FUNCTION_BLOCK FB_Axis EXTENDS FB_Device IMPLEMENTS I_SpeedController
VAR_INPUT
	localEnable		: BOOL; // Enable signal from local Estops, etc. If parent control is configured for enable with no local enable, this can be latched true
	
	{attribute 'OPC.UA.DA' := '1'}
	{attribute 'OPC.UA.DA.StructuredType' := '1'}
	cfg				: ST_AxisConfiguration; 
	
	{attribute 'OPC.UA.DA' := '1'}
	{attribute 'OPC.UA.DA.StructuredType' := '1'}
	ctrlAxis		: ST_AxisControl;
	
	{attribute 'OPC.UA.DA' := '1'} 
	ocmd			: E_AxisCommand;
	
	func			: ST_AxisFunctions;
	
	(* Interlocks/Permissives
	----------------------------------------------------------------------------------------------------*)
	{attribute 'OPC.UA.DA' := '1'}
	{attribute 'OPC.UA.DA.Access' := '1'}
	fwdIntlk		: FB_Permissive;	
	{attribute 'OPC.UA.DA' := '1'}
	{attribute 'OPC.UA.DA.Access' := '1'}
	fwdPerm			: FB_Permissive; 
	{attribute 'OPC.UA.DA' := '1'}
	{attribute 'OPC.UA.DA.Access' := '1'}
	revIntlk		: FB_Permissive; 
	{attribute 'OPC.UA.DA' := '1'}
	{attribute 'OPC.UA.DA.Access' := '1'}
	revPerm			: FB_Permissive; 
	
	(* External inputs
	----------------------------------------------------------------------------------------------------*)
	inpHomeProx AT %I* : BOOL; 				// Link this to home sensor in MapInputs method of Parent
	driveDiagnosticNumber AT %I* : UDINT;	// Link to AX5000 S-0-0390 Diagnostic number
	inpFault		   : BOOL;
	inpFaultText	   : T_MaxString;
END_VAR

VAR_OUTPUT
	{attribute 'OPC.UA.DA' := '1'}
	{attribute 'OPC.UA.DA.StructuredType' := '1'}
	motionParam	: ST_AxisMotionParameters;
	
	{attribute 'OPC.UA.DA' := '1'}
	{attribute 'OPC.UA.DA.Access' := '1'}
	{attribute 'OPC.UA.DA.StructuredType' := '1'}
	sts			: ST_AxisDeviceStatus; 

	{attribute 'OPC.UA.DA' := '1'}
	{attribute 'OPC.UA.DA.Access' := '1'}
	{attribute 'OPC.UA.DA.StructuredType' := '1'}	
	fault		: ST_AxisFault;
END_VAR

VAR PERSISTENT
	offset			: LREAL; // Offset for zero position
	
	{attribute 'OPC.UA.DA' := '1'}
	{attribute 'OPC.UA.DA.Access' := '1'}
	{attribute 'OPC.UA.DA.StructuredType' := '1'}
	positionList	: ARRAY[0..GVL_Lib_ServoConstants.MAX_POSITIONS] OF ST_AxisPosition;
END_VAR

VAR
	axis					: AXIS_REF; 			 // Linked to Motion Axis Object	
	mc						: ST_AxisMotionControl;  // Motion Commands and Parameters
	saveData				: FB_WritePersistentData;
	savePositionListData	: BOOL;	
	resetErrorAndDrive		: BOOL;	
	safeDisable				: BOOL;					 // Disable drive after a safe command, must reset errors to resume operation	
	homingInProgress		: BOOL;					 // Internal bit to set complete flag after homing offset is stored
	mcGearIn				: MC_GearIn;
	mcGearOut				: MC_GearOut;
	
	(* State
	----------------------------------------------------------------------------------------------------*)
	lastGoodState			: E_AxisState;
	nextState				: E_AxisState;
	lastFaultId				: UDINT;
	
	(* Servo Commands
	----------------------------------------------------------------------------------------------------*)
	cmdReceived				: E_AxisCommand;	
	cmdReceivedLast			: E_AxisCommand;	
	pcmd					: E_AxisCommand;	
	pcmdLast				: E_AxisCommand;	
	ocmdLast				: E_AxisCommand;
	storedRelMovePosition	: LREAL;	
	
	(* Speed history/triggers
	----------------------------------------------------------------------------------------------------*)
	jogSpeedLast			: LREAL; 	
	jogSpeedChanged			: BOOL; 	// Jog speed has changed
	ftJogSpeedChanged		: F_TRIG;
	moveSpeedLast			: LREAL;
	moveSpeedChanged		: BOOL;		// Move speed has changed
	ftMoveSpeedChanged		: F_TRIG;
	ftRelMove				: F_TRIG;
	rtAbsMoveADone			: R_TRIG;
	rtAbsMoveBDone			: R_TRIG;
	rtModMoveADone			: R_TRIG;
	rtModMoveBDone			: R_TRIG;

	(* General
	----------------------------------------------------------------------------------------------------*)	
	enableAxisDelay			: TON;
	mcPowerTimeout			: TON;
END_VAR

SUPER^();

Device();
Hmi();
StatusIn();
ProcessCommands();
StateMachine();
MotionControl();
HandleFaults();
StatusOut();
Functions();
SetPositionIds();

METHOD PUBLIC AbsMove
VAR_INPUT
	absMovePosition		: LREAL;
END_VAR
SetMotionParam(param := E_MotorMotionParam.AbsMovePosition, val := absMovePosition);
pcmd := E_AxisCommand.AbsMove;
END_METHOD

METHOD PUBLIC AbsMoveToStoredPosition : BOOL
// Returns true if position is found in list and move started, false otherwise
VAR_INPUT
	id				: INT; 
END_VAR
VAR
	i				: INT;
	success			: BOOL := FALSE;
END_VAR
// Loop through position list to check if the position ID exists and initiate move
FOR i := 0 TO GVL_Lib_ServoConstants.MAX_POSITIONS DO
	// If ID exists in position list
	IF positionList[i].id = id THEN 
		SetMotionParam(param := E_MotorMotionParam.AbsMovePositionId, val := id); // Store commanded position ID
		AbsMove(positionList[i].position); 										  // Initiate absolute move
		success := TRUE;
		EXIT;
	END_IF
END_FOR

AbsMoveToStoredPosition := success;
END_METHOD

METHOD PUBLIC AddFollower
// Must continuously call function
// Execution of coupling or decoupling will be set by 
// the ctrlAxis.coupleFollower bit
VAR_IN_OUT
	follower : AXIS_REF;
END_VAR
IF __ISVALIDREF(follower) THEN
	mcGearIn(Master := axis, Slave := follower, RatioNumerator := cfg.gearRatio, RatioDenominator := 1); 
	mcGearOut(Slave := follower); 

	IF axis.status.homed AND follower.status.homed AND ctrlAxis.coupleFollower
	AND NOT mcGearIn.InGear AND NOT mcGearIn.Execute THEN
		mcGearIn.Execute := TRUE; 
	END_IF

	IF mcGearIn.Execute AND follower.status.coupled THEN 
		mcGearIn.Execute 		:= FALSE;
		ctrlAxis.coupleFollower := TRUE;
	END_IF

	IF mcGearIn.Error THEN
		mcGearIn.Execute := FALSE;
	END_IF

	IF NOT ctrlAxis.coupleFollower AND follower.Status.Coupled THEN 
		mcGearOut.Execute := TRUE;
	END_IF

	IF mcGearOut.Done THEN 
		mcGearOut.Execute := FALSE;
	END_IF

	fault.coupleError 		:= ctrlAxis.coupleFollower AND (NOT axis.Status.Homed OR NOT follower.Status.Homed);
	fault.followerLagError 	:= ctrlAxis.coupleFollower AND axis.Status.Coupled AND follower.Status.Coupled AND
						  	   ABS(axis.NcToPlc.PosDiff - follower.NcToPlc.PosDiff) > cfg.followerLag;			   
END_IF
END_METHOD

METHOD PUBLIC DefinePosition : INT // Check for blank name before overwriting
VAR_INPUT
	id					: INT; // position id
	position			: LREAL; // value of position (mm)
	name				: STRING := ''; // position name
END_VAR
IF positionList[id].name = '' THEN
	DefinePosition := SavePosition(id := id, position := position, name := name);
ELSE
	DefinePosition := 2; // Position has previously been defined. don't overwrite
END_IF
END_METHOD

METHOD PUBLIC DeletePosition : INT
VAR_INPUT
	id : INT;
END_VAR
IF id >= 0 AND id <= GVL_Lib_ServoConstants.MAX_POSITIONS THEN
	positionList[id].name := '';
	positionList[id].position := 0.0;
	DeletePosition := 1; //position deleted, code = 1
ELSE
	DeletePosition := -1; //id out of bounds, code = -1
END_IF
END_METHOD

METHOD PROTECTED Device : BOOL
VAR_INPUT
END_VAR
// to FB device
opTimeout  			 := cfg.opTimeout;
opTimeoutEnable 	 := cfg.opTimeoutEnable;
opActivity 			 := ocmd <> E_AxisCommand.None;

// from FB device
sts.mode	   		 := mode;
sts.modeAuto   		 := sts.mode = E_SystemMode.Auto;
sts.modeManual 		 := sts.mode = E_SystemMode.Manual;
sts.manualOvrde		 := ctrl.manualOvrde; 	
sts.bypass 	   		 := ctrl.bypass;		
sts.sim		   		 := ctrl.sim;			
sts.parentConfigured := parentConfigured;
END_METHOD

METHOD DisableCouple : BOOL
VAR_INPUT
END_VAR
ctrlAxis.coupleFollower := FALSE;
END_METHOD

METHOD PUBLIC DisableLag
pcmd := E_AxisCommand.DisableLag;
END_METHOD

METHOD EnableCouple : BOOL
VAR_INPUT
END_VAR
ctrlAxis.coupleFollower := TRUE;
END_METHOD

METHOD PUBLIC EnableLag
pcmd := E_AxisCommand.EnableLag;
END_METHOD

METHOD PROTECTED Functions
VAR
	i 				: INT;
END_VAR
(* Default function FB calls
----------------------------------------------------------------------------------------------------*)
func.AbsMove(				 	hmiTextStatic := CONCAT(cfg.motorId, ' absolute move'));
func.AbsMoveToStoredPosition(	hmiTextStatic := CONCAT(cfg.motorId, ' absolute move to stored position'));
func.RelMove(					hmiTextStatic := CONCAT(cfg.motorId, ' relative move'));
func.ModMove(				 	hmiTextStatic := CONCAT(cfg.motorId, ' modulus move'));
func.LatchJogFwd(			 	hmiTextStatic := CONCAT(cfg.motorId, ' latch jog forward'));
func.LatchJogRev(				hmiTextStatic := CONCAT(cfg.motorId, ' latch jog reverse'));
func.Home(						hmiTextStatic := CONCAT(cfg.motorId, ' home'));
func.Stop(						hmiTextStatic := CONCAT(cfg.motorId, ' stop'));
func.Couple(					hmiTextStatic := CONCAT(cfg.motorId, ' coupling follower'));
func.Decouple(					hmiTextStatic := CONCAT(cfg.motorId, ' decoupling follower'));
func.ResetDoneBits(				hmiTextStatic := CONCAT(cfg.motorId, ' reset done bits'));

(* Default functions
----------------------------------------------------------------------------------------------------*)

IF func.AbsMove.entry THEN
	FOR i := GVL_Lib_SequencerConstants.MIN_PARAMETERS TO GVL_Lib_SequencerConstants.MAX_PARAMETERS DO
		CASE func.AbsMove.arrParam[i].typeEnum OF
			E_AxisFunctionParam.AbsMovePosition:
				SetMotionParam(param	:= E_MotorMotionParam.AbsMovePosition,
							   val		:= func.AbsMove.arrParam[i].value);
			E_AxisFunctionParam.MoveSpeed:
				SetMotionParam(param	:= E_MotorMotionParam.MoveSpeed,
							   val		:= func.AbsMove.arrParam[i].value);
		END_CASE
	END_FOR
END_IF
IF func.AbsMove.running THEN
	// Check for speed change mid move
	FOR i := GVL_Lib_SequencerConstants.MIN_PARAMETERS TO GVL_Lib_SequencerConstants.MAX_PARAMETERS DO
		IF func.AbsMove.arrParam[i].typeEnum = E_AxisFunctionParam.MoveSpeed THEN
			SetMotionParam(param	:= E_MotorMotionParam.MoveSpeed,
						   val		:= func.AbsMove.arrParam[i].value);
		END_IF
	END_FOR
	// Wait for complete conditions
	func.AbsMove.permComplete.perm.0 S= sts.absMoveComplete;
	
	// Call Action
	IF NOT func.AbsMove.complete AND NOT fault.active
	AND sts.state <> E_AxisState.AbsMove_A AND sts.state <> E_AxisState.AbsMove_B THEN
		// Passing in this motion parameter has the effect of reassigning its own 
		// value to itself. It's done because this input is required for the method
		AbsMove(motionParam.absMovePosition);
	END_IF
	
	func.AbsMove.inpError := fault.active;
END_IF


IF func.AbsMoveToStoredPosition.entry THEN
	FOR i := GVL_Lib_SequencerConstants.MIN_PARAMETERS TO GVL_Lib_SequencerConstants.MAX_PARAMETERS DO
		CASE func.AbsMoveToStoredPosition.arrParam[i].typeEnum OF
			E_AxisFunctionParam.AbsMovePositionId:
				SetMotionParam(param	:= E_MotorMotionParam.AbsMovePositionId,
							   val		:= func.AbsMoveToStoredPosition.arrParam[i].value);
			E_AxisFunctionParam.MoveSpeed:
				SetMotionParam(param	:= E_MotorMotionParam.MoveSpeed,
							   val		:= func.AbsMoveToStoredPosition.arrParam[i].value);
		END_CASE
	END_FOR
END_IF
IF func.AbsMoveToStoredPosition.running THEN
	// Check for speed change mid move
	FOR i := GVL_Lib_SequencerConstants.MIN_PARAMETERS TO GVL_Lib_SequencerConstants.MAX_PARAMETERS DO
		IF func.AbsMoveToStoredPosition.arrParam[i].typeEnum = E_AxisFunctionParam.MoveSpeed THEN
			SetMotionParam(param	:= E_MotorMotionParam.MoveSpeed,
						   val		:= func.AbsMoveToStoredPosition.arrParam[i].value);
		END_IF
	END_FOR
	// Wait for complete conditions
	func.AbsMoveToStoredPosition.permComplete.perm.0 S= sts.absMoveComplete;	
	
	// Call Action
	IF NOT func.AbsMoveToStoredPosition.complete AND NOT fault.active
	AND sts.state <> E_AxisState.AbsMove_A AND sts.state <> E_AxisState.AbsMove_B THEN
		AbsMoveToStoredPosition(motionParam.absMovePositionId);
	END_IF
	
	func.AbsMoveToStoredPosition.inpError := fault.active;
END_IF


IF func.RelMove.entry THEN
	FOR i := GVL_Lib_SequencerConstants.MIN_PARAMETERS TO GVL_Lib_SequencerConstants.MAX_PARAMETERS DO
		CASE func.RelMove.arrParam[i].typeEnum OF
			E_AxisFunctionParam.RelMoveDistance:
				SetMotionParam(param	:= E_MotorMotionParam.RelMoveDistance,
							   val		:= func.RelMove.arrParam[i].value);
			E_AxisFunctionParam.MoveSpeed:
				SetMotionParam(param	:= E_MotorMotionParam.MoveSpeed,
							   val		:= func.RelMove.arrParam[i].value);
		END_CASE
	END_FOR
END_IF
IF func.RelMove.running THEN
	// Check for speed change mid move
	FOR i := GVL_Lib_SequencerConstants.MIN_PARAMETERS TO GVL_Lib_SequencerConstants.MAX_PARAMETERS DO
		IF func.RelMove.arrParam[i].typeEnum = E_AxisFunctionParam.MoveSpeed THEN
			SetMotionParam(param	:= E_MotorMotionParam.MoveSpeed,
						   val		:= func.RelMove.arrParam[i].value);
		END_IF
	END_FOR
	// Wait for complete conditions
	func.RelMove.permComplete.perm.0 S= sts.RelMoveComplete;
	
	// Call Action
	IF NOT func.RelMove.complete AND NOT fault.active
	AND sts.state <> E_AxisState.RelMove_A AND sts.state <> E_AxisState.RelMove_B THEN
		RelMove(motionParam.relMoveDistance);
	END_IF
	
	func.RelMove.inpError := fault.active;
END_IF


IF func.ModMove.entry THEN
	FOR i := GVL_Lib_SequencerConstants.MIN_PARAMETERS TO GVL_Lib_SequencerConstants.MAX_PARAMETERS DO
		CASE func.ModMove.arrParam[i].typeEnum OF
			E_AxisFunctionParam.ModMovePosition:
				SetMotionParam(param	:= E_MotorMotionParam.ModMovePosition,
							   val		:= func.ModMove.arrParam[i].value);
			E_AxisFunctionParam.MoveSpeed:
				SetMotionParam(param	:= E_MotorMotionParam.MoveSpeed,
							   val		:= func.ModMove.arrParam[i].value);
		END_CASE
	END_FOR
	END_IF
IF func.ModMove.running THEN
	// Check for speed change mid move
	FOR i := GVL_Lib_SequencerConstants.MIN_PARAMETERS TO GVL_Lib_SequencerConstants.MAX_PARAMETERS DO
		IF func.ModMove.arrParam[i].typeEnum = E_AxisFunctionParam.MoveSpeed THEN
			SetMotionParam(param	:= E_MotorMotionParam.MoveSpeed,
						   val		:= func.ModMove.arrParam[i].value);
		END_IF
	END_FOR
	// Wait for complete conditions
	func.ModMove.permComplete.perm.0 S= sts.ModMoveComplete;
	
	// Call Action
	IF NOT func.ModMove.complete AND NOT fault.active
	AND sts.state <> E_AxisState.ModMove_A AND sts.state <> E_AxisState.ModMove_B THEN
		ModMove(motionParam.modMovePosition);
	END_IF

	func.ModMove.inpError := fault.active;
END_IF


IF func.LatchJogFwd.entry THEN
	FOR i := GVL_Lib_SequencerConstants.MIN_PARAMETERS TO GVL_Lib_SequencerConstants.MAX_PARAMETERS DO
		CASE func.LatchJogFwd.arrParam[i].typeEnum OF
			E_AxisFunctionParam.JogSpeed: 
				SetMotionParam(param	:= E_MotorMotionParam.JogSpeed,
							   val		:= func.LatchJogFwd.arrParam[i].value);
		END_CASE
	END_FOR
END_IF
IF func.LatchJogFwd.running THEN
	// Check for speed change mid move
	FOR i := GVL_Lib_SequencerConstants.MIN_PARAMETERS TO GVL_Lib_SequencerConstants.MAX_PARAMETERS DO
		IF func.LatchJogFwd.arrParam[i].typeEnum = E_AxisFunctionParam.JogSpeed THEN
			SetMotionParam(param	:= E_MotorMotionParam.JogSpeed,
						   val		:= func.LatchJogFwd.arrParam[i].value);
		END_IF
	END_FOR	
	// Call Action
	IF NOT fault.active THEN
		LatchJogFwd();
	END_IF
	
	// Wait for complete conditions
	func.LatchJogFwd.permComplete.perm.0 S= sts.jogFwdInProgress;
	
	func.LatchJogFwd.inpError := fault.active;
END_IF


IF func.LatchJogRev.entry THEN
	FOR i := GVL_Lib_SequencerConstants.MIN_PARAMETERS TO GVL_Lib_SequencerConstants.MAX_PARAMETERS DO
		CASE func.LatchJogRev.arrParam[i].typeEnum OF
			E_AxisFunctionParam.JogSpeed:
				SetMotionParam(param	:= E_MotorMotionParam.JogSpeed,
							   val		:= func.LatchJogRev.arrParam[i].value);
		END_CASE
	END_FOR
END_IF
IF func.LatchJogRev.running THEN
	// Check for speed change mid move
	FOR i := GVL_Lib_SequencerConstants.MIN_PARAMETERS TO GVL_Lib_SequencerConstants.MAX_PARAMETERS DO
		IF func.LatchJogRev.arrParam[i].typeEnum = E_AxisFunctionParam.JogSpeed THEN
			SetMotionParam(param	:= E_MotorMotionParam.JogSpeed,
						   val		:= func.LatchJogRev.arrParam[i].value);
		END_IF
	END_FOR	
	// Call Action
	IF NOT fault.active THEN
		LatchJogRev();
	END_IF
	
	// Wait for complete conditions
	func.LatchJogRev.permComplete.perm.0 S= sts.jogRevInProgress;
	
	func.LatchJogRev.inpError := fault.active;
END_IF



IF func.Home.entry THEN
	FOR i := GVL_Lib_SequencerConstants.MIN_PARAMETERS TO GVL_Lib_SequencerConstants.MAX_PARAMETERS DO
		CASE func.Home.arrParam[i].typeEnum OF
			E_AxisFunctionParam.HomePosition:
				SetMotionParam(param	:= E_MotorMotionParam.HomePosition,
							   val		:= func.Home.arrParam[i].value);
		END_CASE
	END_FOR
END_IF
IF func.Home.running THEN
	// Wait for complete conditions
	func.Home.permComplete.perm.0 S= sts.homingComplete OR ctrl.sim;
	
	// Call Action
	IF NOT func.Home.complete AND NOT fault.active
	AND sts.state <> E_AxisState.Homing THEN
		Home();
	END_IF
	
	func.Home.inpError := fault.active;
END_IF

IF func.Stop.running THEN
	// Wait for complete conditions	
	func.Stop.permComplete.perm.0 S= sts.stopComplete;
	
	// Call action
	IF NOT func.Stop.complete AND NOT fault.active
	AND sts.state <> E_AxisState.Halting THEN
		Stop();
	END_IF
END_IF


IF func.Couple.running THEN
	ctrlAxis.coupleFollower := TRUE;
	func.Couple.PermComplete.perm.0 := sts.coupled;
END_IF


IF func.Decouple.running THEN
	ctrlAxis.coupleFollower := FALSE;
	func.Decouple.PermComplete.perm.0 := NOT sts.coupled;
END_IF


IF func.ResetDoneBits.running THEN
	ctrlAxis.resetDoneBits := TRUE;
	func.ResetDoneBits.permComplete.perm.0 := TRUE;
END_IF
END_METHOD

METHOD PROTECTED HandleFaults : BOOL
VAR
	i					: INT;
END_VAR
(* ----- Set Faults ----- *)
// Axis Drive Device Error
IF axis.Status.DriveDeviceError THEN
	fault.driveDeviceError := TRUE;
END_IF

// Axis IO Data Invalid
IF axis.Status.IoDataInvalid THEN
	fault.ioDataInvalid := TRUE;
END_IF

// MC_Power Timeout
mcPowerTimeout(IN := (sts.enable AND sts.state > E_AxisState.Power) AND NOT axis.Status.Operational AND NOT resetErrorAndDrive, PT := T#15S);
IF mcPowerTimeout.Q THEN
	fault.mcPowerTimeout := TRUE;
END_IF

// MC_Power Error
IF mc.power.Error THEN
	fault.mcPowerError := TRUE;
END_IF

// MC_MoveVelo Error
IF mc.moveVelocityA.Error OR mc.moveVelocityB.Error THEN
	fault.mcMoveVeloError := TRUE;
END_IF

// MC_MoveAbs Error
IF mc.moveAbsoluteA.Error OR mc.moveAbsoluteB.Error THEN
	fault.mcMoveAbsError := TRUE;
END_IF

// MC_MoveMod Error
IF mc.moveModuloA.Error OR mc.moveModuloB.Error THEN
	fault.mcMoveModError := TRUE;
END_IF

// MC_Halt Command Aborted
IF mc.halt.CommandAborted THEN
	fault.mcHaltCmdAborted := TRUE;
END_IF

// MC_Halt Error
IF mc.halt.Error THEN
	fault.mcHaltError := TRUE;
END_IF

// MC_SetPosition Error
IF mc.setPosition.Error OR mc.readOffset.Error OR mc.writeOffset.Error THEN  //McSetPosition.Error OR
	fault.mcSetPositionError := TRUE;
END_IF

// MC_EnableLag Error
IF mc.enableLag.Error THEN
	fault.mcEnableLagError := TRUE;
END_IF

// MC_DisableLag Error
IF mc.disableLag.Error THEN
	fault.mcDisableLagError := TRUE;
END_IF

// MC_Homing Error
IF mc.homing.Error THEN
	fault.mcHomeError := TRUE;
END_IF

// MC_Reset Error
IF mc.reset.Error THEN
	fault.mcResetError := TRUE;
END_IF

// FB_SoEReset Error
IF mc.resetSoe.Error AND NOT sts.sim THEN
	fault.mcResetSoeError := TRUE;
END_IF

// Other Errors
// (See AddFollower method for more coupling-related errors)
fault.mcGearError := mcGearIn.Error;
fault.external    := inpFault;

(* ----- Handle Reset ----- *)
// The axis will be reset in the upcoming functions call. If that fails, the
// flags will be set high again on the next loop.
IF resetErrorAndDrive THEN
	fault.driveNotOK				:= FALSE;
	fault.driveStateNotOP			:= FALSE;
	fault.driveDeviceError			:= FALSE;
	fault.ioDataInvalid				:= FALSE;
	fault.mcPowerTimeout			:= FALSE;
	fault.mcPowerError				:= FALSE;
	fault.mcMoveVeloError			:= FALSE;
	fault.mcMoveAbsError			:= FALSE;
	fault.mcMoveModError			:= FALSE;
	fault.mcHaltCmdAborted			:= FALSE;
	fault.mcHaltError				:= FALSE;
	fault.mcSetPositionError		:= FALSE;
	fault.mcResetError				:= FALSE;
	fault.mcResetSoeError			:= FALSE;
	fault.mcEnableLagError			:= FALSE;
	fault.mcDisableLagError			:= FALSE;
	fault.mcHomeError				:= FALSE;
	fault.mcGearError				:= FALSE;
	fault.fwdIntlkDisabled 			:= FALSE;
	fault.revIntlkDisabled			:= FALSE;
	fault.coupleError				:= FALSE;
	fault.followerLagError			:= FALSE;
	fault.external					:= FALSE;
	fault.id						:= 0;
	safeDisable						:= FALSE;
	homingInProgress				:= FALSE;
END_IF

IF fault.active THEN
  IF mc.faultId.power <> 0 THEN
	fault.id := mc.faultId.power;
  ELSIF mc.faultId.moveVelocityA <> 0 THEN
	fault.id := mc.faultId.MoveVelocityA;
  ELSIF mc.faultId.moveVelocityB <> 0 THEN
	fault.id := mc.faultId.MoveVelocityB;
  ELSIF mc.faultId.moveAbsoluteA <> 0 THEN
	fault.id := mc.faultId.MoveAbsoluteA;
  ELSIF mc.faultId.moveAbsoluteB <> 0 THEN
	fault.id := mc.faultId.MoveAbsoluteB;
  ELSIF mc.faultId.moveModuloA <> 0 THEN
	fault.id := mc.faultId.MoveModuloA;
  ELSIF mc.faultId.moveModuloB <> 0 THEN
	fault.id := mc.faultId.MoveModuloB;
  ELSIF mc.faultId.halt <> 0 THEN
 	fault.id := mc.faultId.Halt;
  ELSIF mc.faultId.setPosition <> 0 THEN
	fault.id := mc.faultId.SetPosition;
  ELSIF mc.faultId.readOffset <> 0 THEN
	fault.id := mc.faultId.ReadOffset;
  ELSIF mc.faultId.writeOffset <> 0 THEN
	fault.id := mc.faultId.WriteOffset;
  ELSIF mc.faultId.enableLag <> 0 THEN
	fault.id := mc.faultId.EnableLag;
  ELSIF mc.faultId.disableLag <> 0 THEN
	fault.id := mc.faultId.DisableLag;
  ELSIF mc.faultId.homing <> 0 THEN
	fault.id := mc.faultId.Homing;
  ELSIF mc.faultId.reset <> 0 THEN
	fault.id := mc.faultId.Reset;
  ELSIF mc.faultId.resetSoeAds <> 0 AND NOT sts.sim THEN 
	fault.id := mc.faultId.resetSoeAds;
  ELSIF mc.faultId.resetSoeSercos <> 0 THEN
	fault.id := mc.faultId.resetSoeSercos;
  END_IF
  ELSE fault.id := 0; 
END_IF 

// Write message of error on change
IF fault.id = 0 THEN
	fault.ncText := GVL_Lib_TcErrors.List[0].message;
ELSIF lastFaultId <> fault.id THEN
	FOR i := 0 TO GVL_Lib_TcErrors.MAX_INDEX DO
		IF GVL_Lib_TcErrors.List[i].code = fault.id THEN
			fault.ncText := GVL_Lib_TcErrors.List[i].message;
			EXIT;
		END_IF
	END_FOR
END_IF

IF safeDisable THEN // FIXME: Remove once this is configured in our UDT
	IF NOT fwdIntlk.sts.OK AND sts.movingFwd THEN
		fault.inText := CONCAT('Disabled: interlocks lost during motion. fwdIntlk: ', WORD_TO_BINSTR(fwdIntlk.sts.perm, 16));
		fault.fwdIntlkDisabled := TRUE;
	ELSIF NOT revIntlk.sts.OK AND sts.movingRev THEN
		fault.inText := CONCAT('Disabled: interlocks lost during motion. revIntlk: ', WORD_TO_BINSTR(revIntlk.sts.perm, 16));
		fault.revIntlkDisabled := TRUE;
	ELSE
		fault.inText := 'Disabled: external Safe command received.';
	END_IF
ELSIF fault.external THEN
	fault.inText := inpFaultText;
ELSIF fault.mcGearError THEN // FIXME: Remove once this is configured in our UDT
	fault.inText := 'Follower could not be coupled. (Coupling will fail if either axis is moving or faulted for a different reason).';
ELSIF fault.coupleError THEN
	fault.inText := 'Follower could not be coupled. At least one motor was never homed.';
ELSIF fault.followerLagError THEN
	fault.inText := 'Follower lag exceeded the configured threshold';
ELSE
	fault.inText := '';
END_IF

(* ----- Aggregate Faults ----- *)
fault.active := fault.driveNotOK 				OR fault.driveStateNotOP 
				  OR fault.driveDeviceError 	OR fault.ioDataInvalid
				  OR fault.mcPowerTimeout 		OR fault.mcPowerError
				  OR fault.mcMoveVeloError  	OR fault.mcMoveAbsError
				  OR fault.mcMoveModError 		OR fault.mcHomeError
				  OR fault.mcDisableLagError 	OR fault.mcEnableLagError 
				  OR fault.mcHaltCmdAborted 	OR fault.mcHaltError
				  OR fault.mcResetError			OR fault.mcResetSoeError
				  OR fault.mcSetPositionError 	OR safeDisable
				  OR fault.fwdIntlkDisabled		OR fault.revIntlkDisabled
				  OR fault.mcGearError			OR fault.coupleError
				  OR fault.followerLagError		OR fault.external;
END_METHOD

METHOD PROTECTED Hmi
VAR_INPUT
END_VAR
IF ctrlAxis.loadPosition THEN
	ctrlAxis.loadPosition := FALSE;
	LoadPosition(
		id := ctrlAxis.positionToEdit.id,
		position => ctrlAxis.positionToEdit.position,
		name => ctrlAxis.positionToEdit.name
	);
END_IF

IF ctrlAxis.savePosition THEN
	ctrlAxis.savePosition := FALSE;
	SavePosition(
		id := ctrlAxis.positionToEdit.id,
		position := ctrlAxis.positionToEdit.position,
		name := ctrlAxis.positionToEdit.name
	);
END_IF
END_METHOD

METHOD PUBLIC Home
pcmd := E_AxisCommand.Home;
END_METHOD

METHOD PUBLIC JogFwd
pcmd := E_AxisCommand.JogFwd;
END_METHOD

METHOD PUBLIC JogRev
pcmd := E_AxisCommand.JogRev;
END_METHOD

METHOD PUBLIC LatchJogFwd
pcmd := E_AxisCommand.LatchJogFwd;
END_METHOD

METHOD PUBLIC LatchJogRev
pcmd := E_AxisCommand.LatchJogRev;
END_METHOD

METHOD PUBLIC LoadPosition : INT
VAR_INPUT
	id : INT;
END_VAR
VAR_OUTPUT
	position : LREAL;
	name : STRING;
END_VAR
IF id >= 0 AND id <= GVL_Lib_ServoConstants.MAX_POSITIONS THEN
	name := positionList[id].name;
	position := positionList[id].position;
	LoadPosition := 1; //position found, code = 1
ELSE
	LoadPosition := -1; //id out of bounds, code = -1
END_IF
END_METHOD

METHOD PUBLIC ModMove
VAR_INPUT
	modMovePosition		: LREAL;
END_VAR
SetMotionParam(param := E_MotorMotionParam.ModMovePosition, val := modMovePosition);
pcmd := E_AxisCommand.ModMove;
END_METHOD

METHOD PROTECTED MotionControl
VAR
	absMovePos	 : LREAL;
	haltDecel 	 : LREAL;
END_VAR
// Enable the Axis
mc.power(
	Axis				:=	axis, 
	Enable				:=	sts.enable AND sts.state >= E_AxisState.Power,
	Enable_Positive		:=	fwdIntlk.sts.OK, 
	Enable_Negative		:=	revIntlk.sts.OK,
	Override			:=	cfg.powerOverride, 	// 1-100%, 100% typ
	BufferMode			:=	mc.bufferMode, 	 	// MC_Aborting -> Immediate disable; MC_Buffered -> Wait for motion commands to finish before disable
	Status				=>, 
	Busy				=>, 
	Active				=>, 
	Error				=>, 
	ErrorID				=>	mc.faultId.power);

// Move Velocity (A)
mc.moveVelocityA(
	Axis			:=	axis, 
	Execute			:=	(sts.state = E_AxisState.JogFwd_A) 		OR (sts.state = E_AxisState.JogRev_A)
					OR	(sts.state = E_AxisState.LatchJogFwd_A)	OR (sts.state = E_AxisState.LatchJogRev_A), 
	Velocity		:=	motionParam.jogSpeed, 
	Acceleration	:=	motionParam.jogAccel, 
	Deceleration	:=	motionParam.jogDecel, 
	Jerk			:=	motionParam.jerk, 
	Direction		:=	mc.moveDirection, 
	BufferMode		:=	mc.bufferMode, 
	Options			:=	(* Use default values *), 
	InVelocity		=>, 
	Busy			=>, 
	Active			=>, 
	CommandAborted	=>, 
	Error			=>,  
	ErrorID			=>	mc.faultId.moveVelocityA);

// Move Velocity (B)
mc.moveVelocityB(
	Axis			:=	axis, 
	Execute			:=	(sts.state = E_AxisState.JogFwd_B) 		OR (sts.state = E_AxisState.JogRev_B)
					OR	(sts.state = E_AxisState.LatchJogFwd_B) 	OR (sts.state = E_AxisState.LatchJogRev_B), 
	Velocity		:=	motionParam.jogSpeed,    
	Acceleration	:=	motionParam.jogAccel,    
	Deceleration	:=	motionParam.jogDecel,    
	Jerk			:=	motionParam.jerk,    
	Direction		:=	mc.moveDirection, 
	BufferMode		:=	mc.bufferMode,   
	Options			:=	(* Use default values *), 
	InVelocity		=>, 
	Busy			=>, 
	Active			=>, 
	CommandAborted	=>, 
	Error			=>, 
	ErrorID			=>	mc.faultId.moveVelocityB);

// Calculate Move Position (Absolute or Relative)
IF sts.state = E_AxisState.AbsMove_A OR sts.state = E_AxisState.AbsMove_B THEN
	absMovePos := motionParam.absMovePosition;
ELSIF sts.state = E_AxisState.RelMove_A OR sts.state = E_AxisState.RelMove_B THEN
	absMovePos := storedRelMovePosition;
END_IF

// Move Absolute (A)
mc.moveAbsoluteA(
	Axis			:=	axis,
	Execute			:=	sts.state = E_AxisState.AbsMove_A OR sts.state = E_AxisState.RelMove_A,
	Position		:=	absMovePos,
	Velocity		:=	motionParam.moveSpeed,
	Acceleration	:=	motionParam.moveAccel,
	Deceleration	:=	motionParam.moveDecel,
	Jerk			:=	motionParam.jerk,
	BufferMode		:=	mc.bufferMode,
	Options			:=	(* Use default values *),
	Done			=>,
	Busy			=>,
	Active			=>,
	CommandAborted	=>,
	Error			=>, 
	ErrorID			=> mc.faultId.moveAbsoluteA);

// Move Absolute (B)
mc.moveAbsoluteB(
	Axis			:=	axis,
	Execute			:=	sts.state = E_AxisState.AbsMove_B OR sts.state = E_AxisState.RelMove_B,
	Position		:=	absMovePos,
	Velocity		:=	motionParam.moveSpeed,
	Acceleration	:=	motionParam.moveAccel,
	Deceleration	:=	motionParam.moveDecel,
	Jerk			:=	motionParam.jerk,
	BufferMode		:=	mc.bufferMode,
	Options			:=	(* Use default values *),
	Done			=>,
	Busy			=>,
	Active			=>,
	CommandAborted	=>,
	Error			=>, 
	ErrorID			=> mc.faultId.moveAbsoluteB
);

// Move Modulo (A)
mc.moveModuloA(
	Axis			:= axis,
	Execute			:= sts.state = E_AxisState.ModMove_A,
	Position		:= motionParam.modMovePosition,
	Velocity		:= motionParam.moveSpeed,
	Acceleration	:= motionParam.moveAccel,
	Deceleration	:= motionParam.moveDecel,
	Jerk			:= motionParam.jerk,
	Direction		:= MC_Positive_Direction,
	BufferMode		:= mc.bufferMode,
	Options			:=,
	Done			=>,
	Busy			=>,
	Active			=>,
	CommandAborted	=>,
	Error			=>,
	ErrorId			=> mc.faultId.moveModuloA,
	);

// Move Modulo (B)
mc.moveModuloB(
	Axis			:= axis,
	Execute			:= sts.state = E_AxisState.ModMove_B,
	Position		:= motionParam.modMovePosition,
	Velocity		:= motionParam.moveSpeed,
	Acceleration	:= motionParam.moveAccel,
	Deceleration	:= motionParam.moveDecel,
	Jerk			:= motionParam.jerk,
	Direction		:= MC_Positive_Direction,
	BufferMode		:= mc.bufferMode,
	Options			:=,
	Done			=>,      
	Busy			=>,      
	Active			=>,      
	CommandAborted	=>,      
	Error			=>,     
	ErrorId			=> mc.faultId.moveModuloB
	);
	
// Halt
haltDecel := motionParam.haltDecel;
IF haltDecel = 0 THEN
	haltDecel := motionParam.moveDecel;
END_IF
mc.halt(
	Axis			:= axis, 
	Execute			:= sts.state = E_AxisState.Halting  OR sts.state = E_AxisState.Faulting, 
	Deceleration	:= haltDecel, 
	Jerk			:= motionParam.jerk, 
	BufferMode		:= MC_Aborting, 
	Options			:=	(* Use default values *), 
	Done			=>, 
	Busy			=>, 
	Active			=>, 
	CommandAborted	=>, 
	Error			=>,  
	ErrorID			=> mc.faultId.halt);
	
// Teach Position
mc.setPosition(
	Axis			:= axis,
	Execute			:= sts.state = E_AxisState.TeachPositionTemp,
	Position		:= motionParam.teachPosition,
	Mode			:= FALSE,
	Done			=>,
	Busy			=>,
	Error			=>, 
	ErrorID			=> mc.faultId.setPosition);

// Read offset
mc.readOffset(
	Enable 			:= sts.state = E_AxisState.TeachPosition_Read OR sts.state = E_AxisState.InitReadPosition,
	ParameterNumber := AxisEncoderOffset,
	Axis 			:= axis,
	Value 			=>,
	Busy			=>,
	Error			=>, 
	ErrorID			=>	mc.faultId.readOffset);

// Write offset		
mc.writeOffset(
	Execute 		:= sts.state = E_AxisState.TeachPosition_Write OR sts.state = E_AxisState.InitSetPosition,
	ParameterNumber := AxisEncoderOffset,
	Value 			:= offset,
	Axis 			:= axis,
	Busy			=>,
	Error			=>, 
	ErrorID			=> mc.faultId.writeOffset);	
	
// Enable Lag
mc.enableLag(	
	Axis			:= axis,
	Execute			:= sts.state = E_AxisState.EnableLag,
	ParameterNumber := MC_AxisParameter.EnablePosLagMonitoring,
	Value			:= TRUE,
	Done			=>,
	Error			=>,
	ErrorID			=> mc.faultId.enableLag);
	
// Disable Lag
mc.disableLag(	
	Axis			:= axis,
	Execute			:= sts.state = E_AxisState.DisableLag,
	ParameterNumber := MC_AxisParameter.EnablePosLagMonitoring,
	Value			:= FALSE,
	Done			=>,
	Error			=>,
	ErrorID			=> mc.faultId.disableLag);
	
// Homing
mc.homing(
	Axis			:= axis,
	Execute			:= sts.state = E_AxisState.Homing,
	Position		:= motionParam.homePosition,
	HomingMode		:= cfg.homingMode,
	bCalibrationCam	:= inpHomeProx,
	Done			=>,
	Busy			=>,
	Error			=>,
	ErrorId			=> mc.faultId.homing);
	
// Fault Reset
mc.reset(
	Axis		:=	axis, 
	Execute		:=	resetErrorAndDrive OR sts.state = E_AxisState.ResetDrive,
	Done		=>, 
	Busy		=>, 
	Error		=>, 
	ErrorID		=>  mc.faultId.reset);

// Reset - Used for beckhoff servos.
mc.resetSoe(
	NetId		:=	'', 
	Execute		:=	(resetErrorAndDrive OR sts.state = E_AxisState.ResetDrive) AND cfg.isBeckhoffServo AND NOT sts.sim,
	Timeout		:=	T#10S,	// FbSoEReset can take up to 10 seconds 
	Axis		:=	axis, 
	Busy		=>, 
	Error		=>, 
	AdsErrId	=>	, 
	SercosErrId	=>	);
mc.faultId.resetSoeAds 		:= UINT_TO_UDINT(mc.resetSoe.AdsErrId);	
mc.faultId.resetSoeSercos 	:= UINT_TO_UDINT(mc.resetSoe.SercosErrId);

// Read Position
// Used to convert relative move to absolution move
mc.readPosition(
	Enable 			:= TRUE,
	Axis 			:= axis,
	Valid 			=>,
	Busy			=>,
	Error			=>, 
	ErrorID			=>	mc.faultId.readOffset,
	Position		=> );

saveData(
	Port 		:= 851,
	Start 		:= sts.state = E_AxisState.TeachPosition_SaveData OR savePositionListData,
	Mode 		:= SPDM_VAR_BOOST);
	
savePositionListData := FALSE;
END_METHOD

METHOD PROTECTED ProcessCommands
// Check for new valid commands
IF ctrl.reset THEN 
	cmdReceived := E_AxisCommand.Reset;
	ctrl.reset := FALSE;
ELSIF sts.modeManual AND ocmd <> E_AxisCommand.None THEN
	cmdReceived := ocmd;
ELSIF sts.modeAuto AND pcmd <> E_AxisCommand.None THEN
	cmdReceived := pcmd;
END_IF

// Save last commands
IF pcmd <> E_AxisCommand.None THEN
	pcmdLast := pcmd;
END_IF
IF ocmd <> E_AxisCommand.None THEN
	ocmdLast := ocmd;
END_IF
IF cmdReceived <> E_AxisCommand.None THEN
	cmdReceivedLast := cmdReceived;
END_IF

pcmd := E_AxisCommand.None;
ocmd := E_AxisCommand.None;

// Special command handling
resetErrorAndDrive := cmdReceived = E_AxisCommand.Reset;
IF cmdReceived = E_AxisCommand.Safe THEN
	PrvSafe();
END_IF
IF cmdReceived = E_AxisCommand.RelMove AND storedRelMovePosition = 0 THEN
	storedRelMovePosition := sts.position + motionParam.relMoveDistance;
END_IF
IF ftRelMove.Q THEN
	storedRelMovePosition := 0;
END_IF
END_METHOD

METHOD PROTECTED PrvSafe
safeDisable := TRUE;
END_METHOD

METHOD PUBLIC ReadStatus : ST_SpeedControllerStatus
ReadStatus.velocity 	:= sts.velocity;
ReadStatus.torque 		:= sts.torque;
ReadStatus.homed		:= sts.homed;
ReadStatus.coupled 		:= sts.coupled;
ReadStatus.moving 		:= sts.moving;
ReadStatus.movingFwd 	:= sts.movingFwd;
ReadStatus.movingRev 	:= sts.movingRev;
ReadStatus.faulted 		:= fault.active;
END_METHOD

METHOD PUBLIC RelMove
VAR_INPUT
	relMoveDistance		: LREAL;
END_VAR
SetMotionParam(param := E_MotorMotionParam.RelMoveDistance, val := relMoveDistance);
pcmd := E_AxisCommand.RelMove;
END_METHOD

METHOD PUBLIC ResetDoneBits
ctrlAxis.resetDoneBits := TRUE;
END_METHOD

METHOD PUBLIC ResetDrive // Resets drive without resetting errors
pcmd := E_AxisCommand.ResetDrive;
END_METHOD

METHOD PUBLIC Safe
//Command safe regardless of mode
pcmd := E_AxisCommand.Safe;
ocmd := E_AxisCommand.Safe;
END_METHOD

METHOD PUBLIC SavePosition : INT
VAR_INPUT
	id : INT;
	position : LREAL;
	name : STRING;
END_VAR
IF id >= 0 AND id <= GVL_Lib_ServoConstants.MAX_POSITIONS THEN
	positionList[id].name := name;
	positionList[id].position := position;
	SavePosition := 1; //position saved, code = 1
ELSE
	SavePosition := -1; //id out of bounds, code = -1
END_IF
END_METHOD

METHOD PUBLIC SetMotionParam 
VAR_INPUT
	param		: E_MotorMotionParam;
	val			: LREAL;
END_VAR
CASE param OF
	E_MotorMotionParam.JogSpeed:			motionParam.jogSpeed := val;
	E_MotorMotionParam.JogAccel:			motionParam.jogAccel := val;
	E_MotorMotionParam.JogDecel:			motionParam.jogDecel := val;
	E_MotorMotionParam.RelMoveDistance:		motionParam.relMoveDistance := val;
	E_MotorMotionParam.AbsMovePosition:		motionParam.absMovePosition := val;
	E_MotorMotionParam.AbsMovePositionId:	motionParam.absMovePositionId := LREAL_TO_INT(val);
	E_MotorMotionParam.ModMovePosition:		motionParam.modMovePosition := val;
	E_MotorMotionParam.MoveSpeed:			motionParam.moveSpeed := val;
	E_MotorMotionParam.MoveAccel:			motionParam.moveAccel := val;
	E_MotorMotionParam.MoveDecel:			motionParam.moveDecel := val;
	E_MotorMotionParam.Jerk:				motionParam.jerk := val;
	E_MotorMotionParam.TeachPosition:		motionParam.teachPosition := val;
	E_MotorMotionParam.HomePosition:		motionParam.homePosition := val;
	E_MotorMotionParam.HaltDecel:			motionParam.haltDecel := val;
END_CASE
END_METHOD

METHOD INTERNAL SetPositionIds
VAR
	i : INT;
END_VAR
FOR i :=0 TO GVL_Lib_ServoConstants.MAX_POSITIONS DO
	positionList[i].id := i;
END_FOR
END_METHOD

METHOD PROTECTED StateMachine
VAR
	error: INT;
END_VAR
// Reset complete bits
IF NOT cfg.latchDoneBits OR (ctrlAxis.resetDoneBits OR resetErrorAndDrive) THEN
	ctrlAxis.resetDoneBits 		:= FALSE;

	sts.relMoveComplete			:= FALSE;
	sts.absMoveComplete			:= FALSE;
	sts.modMoveComplete			:= FALSE;
	sts.teachPositionComplete	:= FALSE;
	sts.enableLagComplete		:= FALSE;
	sts.disableLagComplete		:= FALSE;
	sts.homingComplete 			:= FALSE;
	sts.resetComplete			:= FALSE;
	sts.stopComplete 			:= FALSE;
END_IF

CASE sts.state OF
		E_AxisState.Off:
			IF sts.enable THEN
				nextState := E_AxisState.InitReadPosition;
			END_IF
			
		E_AxisState.InitReadPosition:
			IF mc.readOffset.Valid THEN
				// check if the offset is already correct
 				IF offset = mc.readOffset.Value THEN
					nextState := E_AxisState.Power;
				ELSE
					nextState := E_AxisState.InitSetPosition;
				END_IF
			END_IF
			
		E_AxisState.InitSetPosition:
			IF mc.writeOffset.Done THEN
				nextState := E_AxisState.InitEnableDelay;
			END_IF
			
		E_AxisState.InitEnableDelay:
			IF enableAxisDelay.Q THEN
				nextState := E_AxisState.Power;
			END_IF
		
		E_AxisState.Power:
			IF sts.enable AND axis.Status.Operational THEN
				nextState := E_AxisState.Enabled;
			END_IF

		E_AxisState.Enabled:
			IF sts.enable AND NOT sts.isFollower THEN				
				IF cmdReceived = E_AxisCommand.JogFwd AND sts.readyFwd THEN
					mc.MoveDirection := MC_Positive_Direction;
					nextState := E_AxisState.JogFwd_A;
				ELSIF cmdReceived = E_AxisCommand.JogRev AND sts.readyRev THEN
					mc.MoveDirection := MC_Negative_Direction;
					nextState := E_AxisState.JogRev_A;
				ELSIF cmdReceived = E_AxisCommand.LatchJogFwd AND sts.readyFwd THEN
					mc.MoveDirection := MC_Positive_Direction;
					nextState := E_AxisState.LatchJogFwd_A;
				ELSIF cmdReceived = E_AxisCommand.LatchJogRev AND sts.readyRev THEN
					mc.MoveDirection := MC_Negative_Direction;
					nextState := E_AxisState.LatchJogRev_A;
				ELSIF cmdReceived = E_AxisCommand.RelMove AND sts.readyRelMove THEN
					nextState := E_AxisState.RelMove_A;
				ELSIF cmdReceived = E_AxisCommand.AbsMove AND sts.readyAbsMove THEN
					nextState := E_AxisState.AbsMove_A;
				ELSIF cmdReceived = E_AxisCommand.ModMove AND sts.readyModMove THEN
					nextState := E_AxisState.ModMove_A;
				ELSIF cmdReceived = E_AxisCommand.TeachPositionTemp THEN
					nextState := E_AxisState.TeachPositionTemp;
				ELSIF cmdReceived = E_AxisCommand.TeachPosition THEN
					nextState := E_AxisState.TeachPosition_Read;
				ELSIF cmdReceived = E_AxisCommand.EnableLag THEN
					nextState := E_AxisState.EnableLag;
				ELSIF cmdReceived = E_AxisCommand.DisableLag THEN
					nextState := E_AxisState.DisableLag;
				ELSIF cmdReceived = E_AxisCommand.Home AND sts.readyFwd AND sts.readyRev THEN
					nextState := E_AxisState.Homing;
				ELSIF cmdReceived = E_AxisCommand.ResetDrive THEN
					nextState := E_AxisState.ResetDrive;
				ELSIF cmdReceived = E_AxisCommand.Stop THEN
					nextState := E_AxisState.Halting;
				END_IF
			END_IF
	
		E_AxisState.JogFwd_A:
			IF cmdReceived <> E_AxisCommand.JogFwd OR mc.moveVelocityA.CommandAborted THEN
				nextState := E_AxisState.Halting;
			ELSIF ftJogSpeedChanged.Q  THEN
				nextState := E_AxisState.JogFwd_B;
			END_IF
			
		E_AxisState.JogFwd_B:
			IF cmdReceived <> E_AxisCommand.JogFwd OR mc.moveVelocityB.CommandAborted THEN
				nextState :=  E_AxisState.Halting;
			ELSIF ftJogSpeedChanged.Q THEN
				nextState := E_AxisState.JogFwd_A;
			END_IF
			
		E_AxisState.JogRev_A:
			IF cmdReceived <> E_AxisCommand.JogRev OR mc.moveVelocityA.CommandAborted THEN
				nextState :=  E_AxisState.Halting;
			ELSIF ftJogSpeedChanged.Q THEN
				nextState := E_AxisState.JogRev_B;
			END_IF
			
		E_AxisState.JogRev_B:
			IF cmdReceived <> E_AxisCommand.JogRev OR mc.moveVelocityB.CommandAborted  THEN
				nextState :=  E_AxisState.Halting;
			ELSIF ftJogSpeedChanged.Q THEN
				nextState := E_AxisState.JogRev_A;
			END_IF	
		
		E_AxisState.LatchJogFwd_A:
			IF cmdReceived = E_AxisCommand.Stop OR mc.moveVelocityA.CommandAborted THEN
				nextState := E_AxisState.Halting;
			ELSIF cmdReceived = E_AxisCommand.LatchJogRev THEN
				IF sts.readyRev THEN
					mc.moveDirection := MC_Negative_Direction;
					nextState := E_AxisState.LatchJogRev_B;
				ELSE
					nextState := E_AxisState.Halting;
				END_IF
			ELSIF ftJogSpeedChanged.Q  THEN
				nextState := E_AxisState.LatchJogFwd_B;
			END_IF
			
		E_AxisState.LatchJogFwd_B:
			IF cmdReceived = E_AxisCommand.Stop OR mc.moveVelocityB.CommandAborted THEN
				nextState :=  E_AxisState.Halting;
			ELSIF cmdReceived = E_AxisCommand.LatchJogRev THEN
				IF sts.readyRev THEN
					mc.moveDirection := MC_Negative_Direction;
					nextState := E_AxisState.LatchJogRev_A;
				ELSE
					nextState := E_AxisState.Halting;
				END_IF
			ELSIF ftJogSpeedChanged.Q THEN
				nextState := E_AxisState.LatchJogFwd_A;
			END_IF
			
		E_AxisState.LatchJogRev_A:	
			IF cmdReceived = E_AxisCommand.Stop OR mc.moveVelocityA.CommandAborted THEN
				nextState :=  E_AxisState.Halting;
			ELSIF cmdReceived = E_AxisCommand.LatchJogFwd THEN
				IF sts.readyFwd THEN
					mc.moveDirection := MC_Positive_Direction;
					nextState := E_AxisState.LatchJogFwd_B;
				ELSE
					nextState := E_AxisState.Halting;
				END_IF
			ELSIF ftJogSpeedChanged.Q THEN
				nextState := E_AxisState.LatchJogRev_B;
			END_IF
			
		E_AxisState.LatchJogRev_B:
			IF cmdReceived = E_AxisCommand.Stop OR mc.moveVelocityB.CommandAborted  THEN
				nextState :=  E_AxisState.Halting;
			ELSIF cmdReceived = E_AxisCommand.LatchJogFwd THEN
				IF sts.readyFwd THEN
					mc.moveDirection := MC_Positive_Direction;
					nextState := E_AxisState.LatchJogFwd_A;
				ELSE
					nextState := E_AxisState.Halting;
				END_IF
			ELSIF ftJogSpeedChanged.Q THEN
				nextState := E_AxisState.LatchJogRev_A;
			END_IF
		
		E_AxisState.RelMove_A:
			IF cmdReceived = E_AxisCommand.Stop THEN
				nextState := E_AxisState.Halting;
			ELSIF ftMoveSpeedChanged.Q THEN
				nextState := E_AxisState.RelMove_B;
			ELSIF rtAbsMoveADone.Q OR mc.MoveAbsoluteA.CommandAborted THEN
				nextState := E_AxisState.Enabled;
				sts.relMoveComplete := TRUE;
			END_IF
			
		E_AxisState.RelMove_B:
			IF cmdReceived = E_AxisCommand.Stop THEN
				nextState := E_AxisState.Halting;
			ELSIF ftMoveSpeedChanged.Q THEN
				nextState := E_AxisState.RelMove_A;
			ELSIF rtAbsMoveBDone.Q OR mc.MoveAbsoluteB.CommandAborted THEN
				nextState := E_AxisState.Enabled;
				sts.relMoveComplete := TRUE;
			END_IF
			
		E_AxisState.AbsMove_A:
			IF cmdReceived = E_AxisCommand.Stop THEN
				nextState := E_AxisState.Halting;
			ELSIF ftMoveSpeedChanged.Q THEN
				nextState := E_AxisState.AbsMove_B;		
			ELSIF rtAbsMoveADone.Q OR mc.MoveAbsoluteA.CommandAborted THEN
				nextState := E_AxisState.Enabled;
				sts.absMoveComplete   := TRUE;
			END_IF
			
		E_AxisState.AbsMove_B:
			IF cmdReceived = E_AxisCommand.Stop THEN
				nextState := E_AxisState.Halting;
			ELSIF ftMoveSpeedChanged.Q THEN
				nextState := E_AxisState.AbsMove_A;
			ELSIF rtAbsMoveBDone.Q OR mc.moveAbsoluteB.CommandAborted THEN
				nextState := E_AxisState.Enabled;
				sts.absMoveComplete   := TRUE;
			END_IF
			
		E_AxisState.ModMove_A:	
			IF cmdReceived = E_AxisCommand.Stop THEN
				nextState := E_AxisState.Halting;
			ELSIF ftMoveSpeedChanged.Q THEN
				nextState := E_AxisState.ModMove_B;		
			ELSIF rtModMoveADone.Q OR mc.moveModuloA.CommandAborted THEN
				nextState := E_AxisState.Enabled;
				sts.modMoveComplete := TRUE;
			END_IF
			
		E_AxisState.ModMove_B:	
			IF cmdReceived = E_AxisCommand.Stop THEN
				nextState := E_AxisState.Halting;
			ELSIF ftMoveSpeedChanged.Q THEN
				nextState := E_AxisState.ModMove_A;		
			ELSIF rtModMoveBDone.Q OR mc.moveModuloB.CommandAborted THEN
				nextState := E_AxisState.Enabled;
				sts.modMoveComplete := TRUE;
			END_IF
			
		E_AxisState.Halting:
			IF mc.halt.Done THEN
				nextState := E_AxisState.Enabled;
				sts.stopComplete := TRUE;
			END_IF
			
		E_AxisState.TeachPositionTemp:  
			IF mc.setPosition.Done THEN
				nextState := E_AxisState.Enabled;
				sts.teachPositionComplete := TRUE;
			END_IF
			
		E_AxisState.TeachPosition_Read: 
			// Read current offset of axis
			IF mc.readOffset.Valid THEN
				offset :=  mc.readOffset.Value + (motionParam.teachPosition - axis.NcToPlc.ActPosWithoutPosCorrection);
				nextState := E_AxisState.TeachPosition_Write;
			END_IF
			
		E_AxisState.TeachPosition_Write: 
			// Write current offset of axis
			IF mc.writeOffset.Done THEN
				nextState := E_AxisState.TeachPosition_SaveData;
			END_IF	
			
		E_AxisState.TeachPosition_SaveData: 
			// Save persistent data to maintain offsets
			IF NOT saveData.BUSY THEN
				nextState := E_AxisState.TeachPosition_EnableDelay;
			END_IF
			
		E_AxisState.TeachPosition_EnableDelay: 
			// Delay while axis is disabled
			IF enableAxisDelay.Q THEN
				nextState := E_AxisState.Power;
				sts.teachPositionComplete := TRUE;
				IF homingInProgress THEN // Indicate homing complete if position was set after homing
					sts.homingComplete := TRUE;
					homingInProgress := FALSE;
				END_IF
			END_IF
		
		E_AxisState.EnableLag:
			IF mc.enableLag.Done THEN
				nextState := E_AxisState.Enabled;
				sts.enableLagComplete	:= TRUE;
			END_IF
			
		E_AxisState.DisableLag:	
			IF mc.disableLag.Done THEN
				nextState := E_AxisState.Enabled;
				sts.disableLagComplete	:= TRUE;
			END_IF
			
		E_AxisState.Homing:	
			homingInProgress := TRUE;	
			IF cmdReceived = E_AxisCommand.Stop THEN
				nextState := E_AxisState.Halting;
			ELSIF mc.homing.Done THEN
				nextState := E_AxisState.TeachPosition_Read;
				SetMotionParam(param := E_MotorMotionParam.TeachPosition, val := axis.NcToPlc.ActPos);
			END_IF
			
		E_AxisState.ResetDrive: 
			IF mc.reset.Done THEN
				nextState := E_AxisState.Enabled;
				sts.resetComplete := TRUE;
			END_IF
			
		E_AxisState.Faulting:
			IF mc.halt.Done OR mc.halt.Error OR mc.halt.CommandAborted THEN
				nextState := E_AxisState.Faulted;
			END_IF	
			
		E_AxisState.Faulted:
			IF NOT fault.active THEN
				nextState := E_AxisState.Off;
			END_IF
END_CASE

// State Transitions from ANY State
IF NOT fault.active AND NOT sts.enable 
AND NOT (sts.state = E_AxisState.Faulting OR sts.state = E_AxisState.Faulted OR sts.state = E_AxisState.Off) THEN
	nextState := E_AxisState.Faulting;
ELSIF fault.active AND NOT (sts.state = E_AxisState.Faulting OR sts.state = E_AxisState.Faulted) THEN
	nextState := E_AxisState.Faulting;
END_IF

sts.state 	:= nextState;
cmdReceived := E_AxisCommand.None;
END_METHOD

METHOD PROTECTED StatusIn
// Axis
axis.ReadStatus(); // Axis status not updated cyclically, must explicitly call
sts.isFollower  := axis.Status.Coupled AND (axis.NcToPlc.CoupleState=3  OR axis.NcToPlc.CoupleState=2); // 1 - Main Motor; 2 - Follower of a Main and Main to a Follower; 3 - Follower only
sts.position	:= axis.NcToPlc.ActPos;
sts.velocity	:= axis.NcToPlc.ActVelo;
sts.torque		:= axis.NcToPlc.ActTorque;
sts.homed       := axis.Status.Homed;
sts.coupled     := axis.NcToPlc.CoupleState<>0;
sts.moving		:= axis.Status.Moving;
sts.movingFwd	:= sts.moving AND sts.velocity > 0;
sts.movingRev	:= sts.moving AND sts.velocity < 0;

sts.enable := localEnable AND NOT safeDisable
			  AND (NOT parentCtrl.estop OR NOT sts.parentConfigured);

// Permissives and Interlocks
fwdIntlk(	bypActive := sts.bypass, cfg := cfg.fwdIntlk);
fwdPerm(	bypActive := sts.bypass, cfg := cfg.fwdPerm);
revIntlk(	bypActive := sts.bypass, cfg := cfg.revIntlk);
revPerm(	bypActive := sts.bypass, cfg := cfg.revPerm);

sts.readyFwd 		:= fwdIntlk.sts.OK AND fwdPerm.sts.OK;
sts.readyRev		:= revIntlk.sts.OK AND revPerm.sts.OK;
sts.readyRelMove	:= sts.state=E_AxisState.Enabled AND
					   ((sts.readyFwd AND (motionParam.relMoveDistance >= 0)) 
					 OR (sts.readyRev AND (motionParam.relMoveDistance <= 0)));
sts.readyAbsMove	:= sts.state=E_AxisState.Enabled AND
					   ((sts.readyFwd AND (motionParam.absMovePosition >= sts.position)) 
					 OR (sts.readyRev AND (motionParam.absMovePosition <= sts.position))); 
sts.readyModMove	:= sts.state=E_AxisState.Enabled AND
					   ((sts.readyFwd AND (motionParam.modMovePosition >= sts.position))  
					 OR (sts.readyRev AND (motionParam.modMovePosition <= sts.position)));

IF sts.moving AND ((NOT fwdIntlk.sts.OK AND sts.movingFwd) OR (NOT revIntlk.sts.OK AND sts.movingRev))
THEN
	PrvSafe();
END_IF

// Timers
enableAxisDelay(IN := sts.state = E_AxisState.InitEnableDelay OR sts.state = E_AxisState.TeachPosition_EnableDelay, PT := cfg.tEnableAxisDelay);

// Check for Speed Change
jogSpeedChanged 			:= motionParam.jogSpeed <> jogSpeedLast;
jogSpeedLast 				:= motionParam.jogSpeed;
ftJogSpeedChanged(CLK		:= jogSpeedChanged);
moveSpeedChanged 			:= motionParam.MoveSpeed <> moveSpeedLast;
moveSpeedLast 				:= motionParam.MoveSpeed;
ftMoveSpeedChanged(CLK		:= moveSpeedChanged);

// Other triggers
ftRelMove(CLK := sts.state = E_AxisState.RelMove_A OR sts.state = E_AxisState.RelMove_B);
rtAbsMoveADone(CLK := mc.moveAbsoluteA.Done);
rtAbsMoveBDone(CLK := mc.moveAbsoluteB.Done);
rtModMoveADone(CLK := mc.moveModuloA.Done);
rtModMoveBDone(CLK := mc.moveModuloB.Done);
END_METHOD

METHOD PROTECTED StatusOut
// Report Command Statuses
sts.jogFwdInProgress 	:= (sts.state = E_AxisState.JogFwd_A 		OR sts.state = E_AxisState.JogFwd_B)
						OR (sts.state = E_AxisState.LatchJogFwd_A 	OR sts.state = E_AxisState.LatchJogFwd_B);
sts.jogRevInProgress 	:= (sts.state = E_AxisState.JogRev_A 		OR sts.state = E_AxisState.JogRev_B)
						OR (sts.state = E_AxisState.LatchJogRev_A	OR sts.state = E_AxisState.LatchJogRev_B);
sts.jogAtSpeed			:= mc.MoveVelocityA.InVelocity OR mc.MoveVelocityB.InVelocity;
sts.relMoveInProgress 	:= (sts.state = E_AxisState.RelMove_A OR sts.state = E_AxisState.RelMove_B);
sts.absMoveInProgress 	:= (sts.state = E_AxisState.AbsMove_A OR sts.state = E_AxisState.AbsMove_B);
sts.modMoveInProgress 	:= (sts.state = E_AxisState.ModMove_A OR sts.state = E_AxisState.ModMove_B);

// Other
sts.driveDiagnosticNumber := driveDiagnosticNumber;
ctrlAxis.resetDoneBits := FALSE;
lastFaultId := fault.id;
IF sts.state < E_AxisState.Faulting THEN
	lastGoodState := sts.state;
END_IF
END_METHOD

METHOD PUBLIC Stop
pcmd := E_AxisCommand.Stop;
END_METHOD

METHOD PUBLIC TeachPosition
VAR_INPUT
	position 		: LREAL;
END_VAR
SetMotionParam(param := E_MotorMotionParam.TeachPosition, val := position);
pcmd := E_AxisCommand.TeachPosition;
END_METHOD

METHOD PUBLIC TeachPositionTemp
VAR_INPUT
	position		: LREAL;
END_VAR
SetMotionParam(param := E_MotorMotionParam.TeachPosition, val := position);
pcmd := E_AxisCommand.TeachPositionTemp;
END_METHOD

END_FUNCTION_BLOCK

(* stored: Version 1.1.0.1, ProductVersion 3.1.4024.12
   POU FB_Axis: Id {e081533c-fdb1-4025-847e-c3bb1b1caa36}, SpecialFunc None
   Folder Protected: Id {930c22f3-10ce-4fd9-b0b4-3631bfb67b16}
   Folder Commands: Id {85a99530-8607-4688-9b94-020d181bfb58}
   Folder Logic: Id {482c5a24-3e6c-41b6-afbc-917e65320721}
   Folder Public: Id {8fca2564-c9b9-4347-b2f7-6e958763f442}
   Folder Commands: Id {4761c3a3-c064-4a6a-97b1-957c9d5db87e}
   Folder Control: Id {17b43a38-ba83-4cf0-be12-706ec11cb865}
   Folder Positions: Id {ff8fd8cd-fa4d-4bda-883b-9d9de0f5559b}
   Method AbsMove: Id {66d48c35-d6eb-45e7-b955-b3cd1dfc4f17}
   Method AbsMoveToStoredPosition: Id {429478c1-e750-4cbe-96b3-37b183561443}
   Method AddFollower: Id {64df873c-d42b-4397-aa9c-62a06db8bdee}
   Method DefinePosition: Id {4efda061-a7e6-46f2-a35d-5b631b4a8a6a}
   Method DeletePosition: Id {4a9bafa8-2bcf-4eaa-a99b-6ceaf7e1193a}
   Method Device: Id {6aaa61cd-4a83-4595-88cd-dc1f255369cf}
   Method DisableCouple: Id {eb58a262-6949-4641-b642-7a8b12b1a2cf}
   Method DisableLag: Id {ad2e7ef3-bd6d-45f2-8417-47a68f3c8be4}
   Method EnableCouple: Id {e2027fcf-f914-4cf5-b84e-6ad552426da1}
   Method EnableLag: Id {5c21c6c7-3917-4ae4-833e-a480bc7faa03}
   Method Functions: Id {c731cb39-62eb-4a45-a95e-13ee5938d5c7}
   Method HandleFaults: Id {cb8fe31f-d608-44af-8f6b-5f5b6d758a4b}
   Method Hmi: Id {3786d032-9989-4ea4-90d7-02874846d9c3}
   Method Home: Id {5e60b3b4-b3b1-463d-9258-f0879e29624a}
   Method JogFwd: Id {e20991aa-f79e-4463-acba-1e069a4912dc}
   Method JogRev: Id {7c2489c3-6e64-476d-b122-12017f403041}
   Method LatchJogFwd: Id {73d51e8e-83b6-49e5-847c-0cd384936e97}
   Method LatchJogRev: Id {e321831d-de3c-4c4c-8da5-3497b45190ac}
   Method LoadPosition: Id {84914dc8-5ad3-4b09-a865-41a50077b9a0}
   Method ModMove: Id {bd416de5-3686-4ccd-8f16-257d39592f28}
   Method MotionControl: Id {99b638d4-42d9-42e0-a7a7-d8379d4e6fa8}
   Method ProcessCommands: Id {2e4561c9-40df-45f1-976c-074e20c2cfd3}
   Method PrvSafe: Id {1c983903-e9ef-46af-95b5-16c3bba4b5ca}
   Method ReadStatus: Id {919179be-6e2f-4b0f-8147-c75ee647ac0b}
   Method RelMove: Id {38878635-83da-4233-a95b-36b6daf62a1f}
   Method ResetDoneBits: Id {6d628401-8689-4c98-9273-cf66471a121c}
   Method ResetDrive: Id {ff4cbb53-89bf-4824-9c00-d86154e102fb}
   Method Safe: Id {4eefb597-de9a-417f-b112-82db1498feff}
   Method SavePosition: Id {c58ec495-30e1-44c0-903b-084e6f794a11}
   Method SetMotionParam: Id {764edde2-1061-44c7-8446-c2c39035b6f5}
   Method SetPositionIds: Id {d2bcda0e-5a33-4031-9ac1-e219c666b520}
   Method StateMachine: Id {82459fb2-7dce-4171-9af9-e02d7052cb8e}
   Method StatusIn: Id {746d9691-1b5a-4806-919d-3fc36431978e}
   Method StatusOut: Id {8fbc8059-4420-4fe0-acda-048d433679b2}
   Method Stop: Id {ad77995b-5b6a-48e4-bfc9-248e43eaf00e}
   Method TeachPosition: Id {ded99c1f-0519-459a-99b2-460f56bb8683}
   Method TeachPositionTemp: Id {5ebeadef-1f86-4668-82c7-33d8ecd1bdeb} *)
